Staubli VAL3: insertIF.pgx

public program insertIF(string x_sKey, num x_nIndex, num& x_nMoveType[], num& x_nIOIndex[], num& x_nValue[], num& x_nANDOR[], bool& x_bToSave)
  local num l_j
  local num l_i
begin
  // insert(trajTemp:tTrajItem[x_sKey].pPointItem[x_nIndex+1])
  append(trajTemp:tTrajItem[x_sKey].pPointItem)

  for l_i = (size(trajTemp:tTrajItem[x_sKey].pPointItem)-1) to(x_nIndex+1) step -1
    // logMsg(toString("",l_i))
    call copyPoint3(x_sKey,l_i,l_i-1)
  endFor
  trajTemp:tTrajItem[x_sKey].pPointItem[x_nIndex+1].pParaItem.nMoveType=8
  for l_i =0 to 2
    trajTemp:tTrajItem[x_sKey].pPointItem[x_nIndex+1].pParaItem.iIfItem.nSigType[l_i]=x_nMoveType[l_i]
    trajTemp:tTrajItem[x_sKey].pPointItem[x_nIndex+1].pParaItem.iIfItem.nSigIndex[l_i]=x_nIOIndex[l_i]
    trajTemp:tTrajItem[x_sKey].pPointItem[x_nIndex+1].pParaItem.iIfItem.nValue[l_i]=x_nValue[l_i]
  endFor
  for l_i = 0 to 1
    trajTemp:tTrajItem[x_sKey].pPointItem[x_nIndex+1].pParaItem.iIfItem.bANDOR[l_i]=(x_nANDOR[l_i]==2)
  endFor

  //trajTemp:libSave()
  x_bToSave=true
end
